(* PLC project Vn_op_mux, Beckhoff Automation GmbH TwinCAT PLC Control 3.5.13.21 *)
(* stored: creationDateTime 1970-01-01T00:00:00 *)

PROGRAM Vn_op_mux

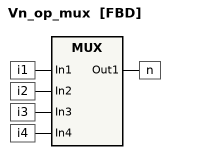
(* FBD diagram, written out as Structured Text *)
n := MUX(i1, i2, i3, i4);
END_PROGRAM
